FUNCTION_BLOCK FB_ClientSendMsg
(*

The function block used to send cyclic message strings.

Basie on orginal Beckhoffs example.

Constructor: 	Patryk Panylo
Company:		E. Riexinger GmbH
Date:			18.02.2019
Version:		1.00

Date:			Revision:		Who:				Comment
dd.mm.yyyy		x.xx			Initials			comment

*)
VAR_INPUT
	(* Input variables / Eingang Variablen *)
	bEnable						:BOOL;					(* Enable FB *)
	bExecute					:BOOL := FALSE;			(* Send string *)
	sMsg						:T_MaxString := '';
	sPrefix						:STRING := '';			(* Message prefix *)
	sSuffix						:STRING := '';			(* Message suffix *)
END_VAR
VAR_OUTPUT
	(* Output variables / Ausgang Variablen *)
	bErrorSndFifoOverflow 		:BOOL := FALSE;			(* Send fifo overflow error *)
END_VAR
VAR_IN_OUT
	(* Input Output variables / Ausgang Variablen *)
	fbTx 						:FB_FrameFifo;			(* Tx fifo *)
	fbLoggger					:FB_LogFifo;			(* Logger message fifo *)
	arsMsg						:ARRAY[1..GVL_TCPIP.RECEIVE_MESSAGE_MAX] OF T_MaxString;			(* Get message of received an ASCII typable string data. *)
END_VAR
VAR
	(* Enummerations *)
	
	(* Variables *)
	
	(* References *)

	(* Interfaces *)

	(* Instances *)
	rtExecute					:R_TRIG;
END_VAR


IF NOT bEnable
THEN
	RETURN;
END_IF

rtExecute(CLK := bExecute);
bErrorSndFifoOverflow := FALSE;
IF rtExecute.Q
THEN
	(* Put string to the tx fifo *)
	fbTx.AddTail(			
		sPut := CONCAT(CONCAT(sPrefix, sMsg), sSuffix)
	);
	
	MEMSET(ADR(arsMsg),0,SIZEOF(arsMsg));												(* Clear Rx frame *)
	
	IF NOT fbTx.bOk (* TX fifo overflow => log error *)
	THEN
		fbLoggger.Error(
			sMessage := 'FB_FrameFifo(sender)', 
			nErrID := GVL_TCPIP.ERROR_SENDFIFO_OVERFLOW 
		);
		
		bErrorSndFifoOverflow := TRUE;
	END_IF

END_IF

END_FUNCTION_BLOCK

(* stored: Version 1.1.0.1, ProductVersion 3.1.4024.15
   POU FB_ClientSendMsg: Id {09c10c50-b482-4c06-b5b0-de3cc0e5479b}, SpecialFunc None *)
